(* IEC 61131-3 sources: trust-platform/editors/vscode/media/examples/conveyor/src, 2 files *)

(* ---- Configuration.st ---- *)
CONFIGURATION ConveyorCell
TASK Cycle (INTERVAL := T#50ms, PRIORITY := 1);
PROGRAM P1 WITH Cycle : MainProgram;
VAR_CONFIG
    P1.e_stop         AT %IX0.0 : BOOL;
    P1.running        AT %QX2.0 : BOOL;
    P1.conveyor_speed AT %QW0   : INT;
    P1.part_count     AT %MW0   : INT;
END_VAR
END_CONFIGURATION

(* ---- Main.st ---- *)
PROGRAM MainProgram
VAR
    e_stop         : BOOL;   (* %IX0.0 — write TRUE to stop the line *)
    running        : BOOL;   (* %QX2.0 *)
    conveyor_speed : INT;    (* %QW0   *)
    part_count     : INT;    (* %MW0   *)
END_VAR

running := NOT e_stop;
IF running THEN
    IF conveyor_speed < 100 THEN
        conveyor_speed := conveyor_speed + 5;
    ELSE
        part_count := part_count + 1;
        conveyor_speed := 0;
    END_IF;
ELSE
    conveyor_speed := 0;
END_IF;
END_PROGRAM
